// Characterization of FB_MonetTelescopeControl for a park or a stop that arrives during the power-on, and for an Init() during a
// park, on mock axes (plan step 1, MONETcommonTests README). These tests pin what the code does today, with the line of the
// behaviour in a comment; they are not a specification. Every test owns a rig and runs over many PLC cycles (VAR_INST of the
// method, one Scan() per cycle). Failed checks are also noted in GVL_Diag.sFailures (printed by Run-Tests.ps1).
FUNCTION_BLOCK MonetParkDuringPowerOn_Tests EXTENDS TcUnit.FB_TestSuite
VAR
END_VAR

Park_During_PowerOn_Parks_In_Place_And_Closes_The_Covers();
Park_During_Homing_Stops_The_Homing_Axes_First();
Stop_During_PowerOn_Aborts_The_Startup();
Init_During_Park_Is_Refused();
Startup_Finished_Is_Logged_At_The_Completion();
Stop_During_The_Move_To_Home_Logs_No_Startup_Finished();

// M:533-545 (#87), M:1245 (#113): a park that arrives while the power-on has only commanded the covers aborts the power-on and
// parks in place (no axis is calibrated, so none is sent to the park position): the axes are disabled, the covers that the
// power-on opened are closed again, READY_STATE is parked (0.0).
METHOD PRIVATE Park_During_PowerOn_Parks_In_Place_And_Closes_The_Covers
VAR_INST
	rig			: FB_MonetRig;
	nStep		: INT;
	nCycles		: UINT;
	sTest		: STRING(80);
END_VAR
TEST('Park_During_PowerOn_Parks_In_Place_And_Closes_The_Covers');
sTest := 'Park_During_PowerOn_Parks_In_Place_And_Closes_The_Covers: ';
IF nStep >= 90 THEN
	RETURN;
END_IF
rig.Scan();
nCycles := nCycles + 1;
CASE nStep OF
0:	// wait for the clock, then power on
	IF rig.ClockValid THEN
		rig.fbTel.Init();
		nStep := 10;
		nCycles := 0;
	ELSIF nCycles > 2000 THEN
		AssertTrue(Condition := FALSE, Message := 'the astronomical clock never became valid');
		F_Note(bFailed := TRUE, sText := CONCAT(sTest, 'the astronomical clock never became valid'));
		nStep := 99;
		TEST_FINISHED();
	END_IF
10:	// the power-on has commanded the covers: park now
	IF rig.fbCovers.nOpenCalls >= 1 THEN
		rig.fbTel.Park();
		nStep := 20;
		nCycles := 0;
	ELSIF nCycles > 300 THEN
		AssertTrue(Condition := FALSE, Message := 'the power-on never commanded the covers');
		F_Note(bFailed := TRUE, sText := CONCAT(sTest, 'the power-on never commanded the covers'));
		nStep := 99;
		TEST_FINISHED();
	END_IF
20:	// wait until the park has finished
	IF rig.fbTel.bIsParked AND nCycles > 5 THEN
		AssertFalse(Condition := rig.fbTel.bParkActive, Message := 'the park is over');
		F_Note(bFailed := (rig.fbTel.bParkActive), sText := CONCAT(sTest, 'the park is over'));
		AssertTrue(Condition := rig.fbCovers.bClosed AND rig.fbCovers.nCloseCalls >= 1, Message := 'the covers the power-on opened are closed again');
		F_Note(bFailed := NOT (rig.fbCovers.bClosed AND rig.fbCovers.nCloseCalls >= 1), sText := CONCAT(sTest, 'the covers the power-on opened are closed again'));
		AssertFalse(Condition := rig.fbElev.bEnable OR rig.fbAzim.bEnable OR rig.fbDero.bEnable, Message := 'all three axes are disabled (parked in place)');
		F_Note(bFailed := (rig.fbElev.bEnable OR rig.fbAzim.bEnable OR rig.fbDero.bEnable), sText := CONCAT(sTest, 'all three axes are disabled (parked in place)'));
		AssertTrue(Condition := rig.fbElev.nStopEdges = 0 AND rig.fbAzim.nStopEdges = 0 AND rig.fbDero.nStopEdges = 0, Message := 'nothing was moving, so no axis was stopped');
		F_Note(bFailed := NOT (rig.fbElev.nStopEdges = 0 AND rig.fbAzim.nStopEdges = 0 AND rig.fbDero.nStopEdges = 0), sText := CONCAT(sTest, 'nothing was moving, so no axis was stopped'));
		AssertFalse(Condition := rig.fbTel.fbStartup.Initializing, Message := 'the startup is aborted');
		F_Note(bFailed := (rig.fbTel.fbStartup.Initializing), sText := CONCAT(sTest, 'the startup is aborted'));
		AssertTrue(Condition := rig.fbTel.ReadyState = 0.0, Message := 'READY_STATE is parked (0.0)');
		F_Note(bFailed := NOT (rig.fbTel.ReadyState = 0.0), sText := CONCAT(sTest, 'READY_STATE is parked (0.0)'));
		nStep := 99;
		TEST_FINISHED();
	ELSIF nCycles > 600 THEN
		AssertTrue(Condition := FALSE, Message := 'the park did not finish');
		F_Note(bFailed := TRUE, sText := CONCAT(sTest, 'the park did not finish'));
		nStep := 99;
		TEST_FINISHED();
	END_IF
END_CASE
END_METHOD

// M:533-545 (#87) with the abort stop (#84): a park that arrives while the axes are homing aborts the power-on, sends one stop to
// each axis that was homing, waits for the stop to settle and then parks in place; the aborted homing does not calibrate.
METHOD PRIVATE Park_During_Homing_Stops_The_Homing_Axes_First
VAR_INST
	rig			: FB_MonetRig;
	nStep		: INT;
	nCycles		: UINT;
	sTest		: STRING(80);
END_VAR
TEST('Park_During_Homing_Stops_The_Homing_Axes_First');
sTest := 'Park_During_Homing_Stops_The_Homing_Axes_First: ';
IF nStep >= 90 THEN
	RETURN;
END_IF
rig.Scan();
nCycles := nCycles + 1;
CASE nStep OF
0:	// wait for the clock, then power on
	IF rig.ClockValid THEN
		rig.SetHomeScans(40);
		rig.fbTel.Init();
		nStep := 10;
		nCycles := 0;
	ELSIF nCycles > 2000 THEN
		AssertTrue(Condition := FALSE, Message := 'the astronomical clock never became valid');
		F_Note(bFailed := TRUE, sText := CONCAT(sTest, 'the astronomical clock never became valid'));
		nStep := 99;
		TEST_FINISHED();
	END_IF
10:	// both axes are homing: park now
	IF rig.fbElev.fbAxis.Homing AND rig.fbAzim.fbAxis.Homing THEN
		rig.fbTel.Park();
		nStep := 20;
		nCycles := 0;
	ELSIF nCycles > 300 THEN
		AssertTrue(Condition := FALSE, Message := 'the axes never started homing');
		F_Note(bFailed := TRUE, sText := CONCAT(sTest, 'the axes never started homing'));
		nStep := 99;
		TEST_FINISHED();
	END_IF
20:	// wait until the park has finished
	IF rig.fbTel.bIsParked AND nCycles > 5 THEN
		AssertTrue(Condition := rig.fbElev.nStopEdges = 1 AND rig.fbAzim.nStopEdges = 1, Message := 'the elevation and the azimuth that were homing got one stop each');
		F_Note(bFailed := NOT (rig.fbElev.nStopEdges = 1 AND rig.fbAzim.nStopEdges = 1), sText := CONCAT(sTest, 'the elevation and the azimuth that were homing got one stop each'));
		AssertFalse(Condition := rig.fbElev.Calibrated OR rig.fbAzim.Calibrated, Message := 'the aborted homing did not calibrate');
		F_Note(bFailed := (rig.fbElev.Calibrated OR rig.fbAzim.Calibrated), sText := CONCAT(sTest, 'the aborted homing did not calibrate'));
		AssertFalse(Condition := rig.fbElev.bEnable OR rig.fbAzim.bEnable OR rig.fbDero.bEnable, Message := 'all three axes are disabled (parked in place)');
		F_Note(bFailed := (rig.fbElev.bEnable OR rig.fbAzim.bEnable OR rig.fbDero.bEnable), sText := CONCAT(sTest, 'all three axes are disabled (parked in place)'));
		AssertTrue(Condition := rig.fbCovers.bClosed, Message := 'the covers are closed');
		F_Note(bFailed := NOT (rig.fbCovers.bClosed), sText := CONCAT(sTest, 'the covers are closed'));
		AssertTrue(Condition := rig.fbTel.ReadyState = 0.0, Message := 'READY_STATE is parked (0.0)');
		F_Note(bFailed := NOT (rig.fbTel.ReadyState = 0.0), sText := CONCAT(sTest, 'READY_STATE is parked (0.0)'));
		nStep := 99;
		TEST_FINISHED();
	ELSIF nCycles > 800 THEN
		AssertTrue(Condition := FALSE, Message := 'the park did not finish');
		F_Note(bFailed := TRUE, sText := CONCAT(sTest, 'the park did not finish'));
		nStep := 99;
		TEST_FINISHED();
	END_IF
END_CASE
END_METHOD

// M:508-518 (#80): a stop outranks a running power-on. The startup is aborted (READY_STATE -2.0), nothing is parked, and the
// covers the power-on opened stay open: a stop does not close them.
METHOD PRIVATE Stop_During_PowerOn_Aborts_The_Startup
VAR_INST
	rig			: FB_MonetRig;
	nStep		: INT;
	nCycles		: UINT;
	sTest		: STRING(80);
END_VAR
TEST('Stop_During_PowerOn_Aborts_The_Startup');
sTest := 'Stop_During_PowerOn_Aborts_The_Startup: ';
IF nStep >= 90 THEN
	RETURN;
END_IF
rig.Scan();
nCycles := nCycles + 1;
CASE nStep OF
0:	// wait for the clock, then power on
	IF rig.ClockValid THEN
		rig.fbTel.Init();
		nStep := 10;
		nCycles := 0;
	ELSIF nCycles > 2000 THEN
		AssertTrue(Condition := FALSE, Message := 'the astronomical clock never became valid');
		F_Note(bFailed := TRUE, sText := CONCAT(sTest, 'the astronomical clock never became valid'));
		nStep := 99;
		TEST_FINISHED();
	END_IF
10:	// the power-on has commanded the covers: stop now
	IF rig.fbCovers.nOpenCalls >= 1 THEN
		rig.fbTel.Stop();
		nStep := 20;
		nCycles := 0;
	ELSIF nCycles > 300 THEN
		AssertTrue(Condition := FALSE, Message := 'the power-on never commanded the covers');
		F_Note(bFailed := TRUE, sText := CONCAT(sTest, 'the power-on never commanded the covers'));
		nStep := 99;
		TEST_FINISHED();
	END_IF
20:	// wait until the stop has settled
	IF NOT rig.fbTel.bStopActive AND rig.fbTel.bStopped AND nCycles > 5 THEN
		AssertFalse(Condition := rig.fbTel.bPowerActive, Message := 'the power-on request is dropped');
		F_Note(bFailed := (rig.fbTel.bPowerActive), sText := CONCAT(sTest, 'the power-on request is dropped'));
		AssertFalse(Condition := rig.fbTel.bParkActive OR rig.fbTel.bIsParked, Message := 'the stop does not park');
		F_Note(bFailed := (rig.fbTel.bParkActive OR rig.fbTel.bIsParked), sText := CONCAT(sTest, 'the stop does not park'));
		AssertTrue(Condition := rig.fbTel.ReadyState = -2.0, Message := 'READY_STATE is -2.0 (startup aborted)');
		F_Note(bFailed := NOT (rig.fbTel.ReadyState = -2.0), sText := CONCAT(sTest, 'READY_STATE is -2.0 (startup aborted)'));
		AssertTrue(Condition := rig.fbCovers.bOpened, Message := 'the covers stay open');
		F_Note(bFailed := NOT (rig.fbCovers.bOpened), sText := CONCAT(sTest, 'the covers stay open'));
		nStep := 99;
		TEST_FINISHED();
	ELSIF nCycles > 400 THEN
		AssertTrue(Condition := FALSE, Message := 'the stop did not settle');
		F_Note(bFailed := TRUE, sText := CONCAT(sTest, 'the stop did not settle'));
		nStep := 99;
		TEST_FINISHED();
	END_IF
END_CASE
END_METHOD

// M:1969 (#87, #80): park wins in both orders. An Init() while a park runs is refused with a reason and starts no power-on; the
// park goes on and ends parked.
METHOD PRIVATE Init_During_Park_Is_Refused
VAR_INST
	rig			: FB_MonetRig;
	nStep		: INT;
	nCycles		: UINT;
	sTest		: STRING(80);
END_VAR
TEST('Init_During_Park_Is_Refused');
sTest := 'Init_During_Park_Is_Refused: ';
IF nStep >= 90 THEN
	RETURN;
END_IF
rig.Scan();
nCycles := nCycles + 1;
CASE nStep OF
0:	// wait for the clock, then power on
	IF rig.ClockValid THEN
		rig.fbTel.Init();
		nStep := 10;
		nCycles := 0;
	ELSIF nCycles > 2000 THEN
		AssertTrue(Condition := FALSE, Message := 'the astronomical clock never became valid');
		F_Note(bFailed := TRUE, sText := CONCAT(sTest, 'the astronomical clock never became valid'));
		nStep := 99;
		TEST_FINISHED();
	END_IF
10:	// online: start a park
	IF rig.Online THEN
		rig.fbTel.Park();
		nStep := 20;
		nCycles := 0;
	ELSIF nCycles > 1500 THEN
		AssertTrue(Condition := FALSE, Message := 'the mock telescope did not reach READY_STATE 1.0');
		F_Note(bFailed := TRUE, sText := CONCAT(sTest, 'the mock telescope did not reach READY_STATE 1.0'));
		nStep := 99;
		TEST_FINISHED();
	END_IF
20:	// the park is running: an Init() now is refused
	rig.fbTel.Init();
		AssertTrue(Condition := rig.fbTel.bInitRefused, Message := 'the Init() is refused');
		F_Note(bFailed := NOT (rig.fbTel.bInitRefused), sText := CONCAT(sTest, 'the Init() is refused'));
		AssertTrue(Condition := rig.fbTel.sInitRefusedReason = 'park in progress, send stop to cancel it', Message := 'the reason names the park');
		F_Note(bFailed := NOT (rig.fbTel.sInitRefusedReason = 'park in progress, send stop to cancel it'), sText := CONCAT(sTest, 'the reason names the park'));
		AssertFalse(Condition := rig.fbTel.bPowerActive, Message := 'no power-on is started');
		F_Note(bFailed := (rig.fbTel.bPowerActive), sText := CONCAT(sTest, 'no power-on is started'));
	nStep := 30;
	nCycles := 0;
30:	// wait until the park has finished
	IF rig.fbTel.bIsParked AND nCycles > 5 THEN
		AssertFalse(Condition := rig.fbTel.bPowerActive, Message := 'the power-on request is still dropped');
		F_Note(bFailed := (rig.fbTel.bPowerActive), sText := CONCAT(sTest, 'the power-on request is still dropped'));
		AssertTrue(Condition := rig.fbTel.ReadyState = 0.0, Message := 'the park ended parked (0.0)');
		F_Note(bFailed := NOT (rig.fbTel.ReadyState = 0.0), sText := CONCAT(sTest, 'the park ended parked (0.0)'));
		nStep := 99;
		TEST_FINISHED();
	ELSIF nCycles > 800 THEN
		AssertTrue(Condition := FALSE, Message := 'the park did not finish');
		F_Note(bFailed := TRUE, sText := CONCAT(sTest, 'the park did not finish'));
		nStep := 99;
		TEST_FINISHED();
	END_IF
END_CASE
END_METHOD

// #287: 'startup finished' is logged when the power-on completes (stage complete), not when the axes are ready at the
// start of the move to home.
METHOD PRIVATE Startup_Finished_Is_Logged_At_The_Completion
VAR_INST
	rig			: FB_MonetRig;
	nStep		: INT;
	nCycles		: UINT;
	sTest		: STRING(80);
	bSawMove	: BOOL;
	bEarly		: BOOL;
END_VAR
TEST('Startup_Finished_Is_Logged_At_The_Completion');
sTest := 'Startup_Finished_Is_Logged_At_The_Completion: ';
IF nStep >= 90 THEN
	RETURN;
END_IF
IF nStep = 0 AND nCycles = 0 THEN
	rig.WatchLog(sText := 'startup finished');
END_IF
rig.Scan();
nCycles := nCycles + 1;
CASE nStep OF
0:	// wait for the clock, then power on
	IF rig.ClockValid THEN
		rig.fbTel.Init();
		nStep := 10;
		nCycles := 0;
	ELSIF nCycles > 2000 THEN
		AssertTrue(Condition := FALSE, Message := 'the astronomical clock never became valid');
		F_Note(bFailed := TRUE, sText := CONCAT(sTest, 'the astronomical clock never became valid'));
		nStep := 99;
		TEST_FINISHED();
	END_IF
10:	// the move to home: no 'startup finished' yet
	IF rig.fbTel.ePowerOnStage = E_PowerOnStage.wait_home THEN
		bSawMove := TRUE;
		IF rig.LogHits > 0 THEN
			bEarly := TRUE;
		END_IF
	END_IF
	IF rig.Online THEN
		nStep := 20;
		nCycles := 0;
	ELSIF nCycles > 1500 THEN
		AssertTrue(Condition := FALSE, Message := 'the mock telescope did not reach READY_STATE 1.0');
		F_Note(bFailed := TRUE, sText := CONCAT(sTest, 'the mock telescope did not reach READY_STATE 1.0'));
		nStep := 99;
		TEST_FINISHED();
	END_IF
20:	// a few scans after the completion: logged once
	IF nCycles >= 5 THEN
		AssertTrue(Condition := bSawMove, Message := 'the power-on moved to home');
		F_Note(bFailed := NOT (bSawMove), sText := CONCAT(sTest, 'the power-on moved to home'));
		AssertTrue(Condition := NOT bEarly, Message := 'no startup finished during the move to home');
		F_Note(bFailed := NOT (NOT bEarly), sText := CONCAT(sTest, 'no startup finished during the move to home'));
		AssertTrue(Condition := rig.LogHits = 1, Message := 'startup finished is logged once at the completion');
		F_Note(bFailed := NOT (rig.LogHits = 1), sText := CONCAT(sTest, 'startup finished is logged once at the completion'));
		nStep := 99;
		TEST_FINISHED();
	END_IF
END_CASE
END_METHOD

// #287: a power-on stopped during the move to home never logs 'startup finished' (MONET/N 2026-11-13: it did, at the start
// of the move).
METHOD PRIVATE Stop_During_The_Move_To_Home_Logs_No_Startup_Finished
VAR_INST
	rig			: FB_MonetRig;
	nStep		: INT;
	nCycles		: UINT;
	sTest		: STRING(80);
	nInMove		: UINT;
END_VAR
TEST('Stop_During_The_Move_To_Home_Logs_No_Startup_Finished');
sTest := 'Stop_During_The_Move_To_Home_Logs_No_Startup_Finished: ';
IF nStep >= 90 THEN
	RETURN;
END_IF
IF nStep = 0 AND nCycles = 0 THEN
	rig.WatchLog(sText := 'startup finished');
END_IF
rig.Scan();
nCycles := nCycles + 1;
CASE nStep OF
0:	// wait for the clock, then power on
	IF rig.ClockValid THEN
		rig.fbTel.Init();
		nStep := 10;
		nCycles := 0;
	ELSIF nCycles > 2000 THEN
		AssertTrue(Condition := FALSE, Message := 'the astronomical clock never became valid');
		F_Note(bFailed := TRUE, sText := CONCAT(sTest, 'the astronomical clock never became valid'));
		nStep := 99;
		TEST_FINISHED();
	END_IF
10:	// stop during the move to home
	IF rig.fbTel.ePowerOnStage = E_PowerOnStage.wait_home AND rig.fbElev.MoveAxis THEN
		nInMove := nInMove + 1;
	END_IF
	IF nInMove >= 5 THEN
		rig.fbTel.Stop();
		nStep := 20;
		nCycles := 0;
	ELSIF nCycles > 1500 THEN
		AssertTrue(Condition := FALSE, Message := 'the power-on did not move to home');
		F_Note(bFailed := TRUE, sText := CONCAT(sTest, 'the power-on did not move to home'));
		nStep := 99;
		TEST_FINISHED();
	END_IF
20:	// the stop has settled: the power-on is aborted and nothing claims a finished startup
	IF NOT rig.fbTel.bStopActive AND rig.fbTel.bStopped AND nCycles > 20 THEN
		AssertTrue(Condition := NOT rig.fbTel.bPowerActive AND rig.fbTel.ReadyState = -2.0, Message := 'the power-on is aborted (READY_STATE -2.0)');
		F_Note(bFailed := NOT (NOT rig.fbTel.bPowerActive AND rig.fbTel.ReadyState = -2.0), sText := CONCAT(sTest, 'the power-on is aborted (READY_STATE -2.0)'));
		AssertTrue(Condition := rig.LogHits = 0, Message := 'no startup finished for a stopped power-on');
		F_Note(bFailed := NOT (rig.LogHits = 0), sText := CONCAT(sTest, 'no startup finished for a stopped power-on'));
		nStep := 99;
		TEST_FINISHED();
	ELSIF nCycles > 400 THEN
		AssertTrue(Condition := FALSE, Message := 'the stop did not settle');
		F_Note(bFailed := TRUE, sText := CONCAT(sTest, 'the stop did not settle'));
		nStep := 99;
		TEST_FINISHED();
	END_IF
END_CASE
END_METHOD

END_FUNCTION_BLOCK

(* stored: Version 1.1.0.1, ProductVersion 3.1.4024.15
   POU MonetParkDuringPowerOn_Tests: Id {ef273f8d-20bc-4a45-b4f7-010fd9017fa8}, SpecialFunc None
   Method Park_During_PowerOn_Parks_In_Place_And_Closes_The_Covers: Id {27f535d0-bbf6-4f9b-b4ca-266f7b7d2542}
   Method Park_During_Homing_Stops_The_Homing_Axes_First: Id {71651cc9-a542-4aa6-9cd5-b52ae8699fee}
   Method Stop_During_PowerOn_Aborts_The_Startup: Id {25600afc-21e9-4323-b67d-f3e061c4061a}
   Method Init_During_Park_Is_Refused: Id {106ad422-b016-4cc5-b9f2-4d1c7175e978}
   Method Startup_Finished_Is_Logged_At_The_Completion: Id {7fcc7d61-3643-47a4-b9b5-587334bfdbca}
   Method Stop_During_The_Move_To_Home_Logs_No_Startup_Finished: Id {987a80d1-3fa0-45b3-afa0-c6ac188f6d16} *)
